{attribute 'qualified_only'}
VAR_GLOBAL
    fbPersistentDataStorage : LCLS_Tc_DevAbs.FB_PersistentDataStorage;
    eModeSelect : E_ModeSelector := E_ModeSelector.ModeNone;
END_VAR

(* stored: Version 1.1.0.1
   GVL GVL_Common: Id {327df3f0-49dd-4578-a690-f7d367af622c} *)
